(* IEC 61131-3 sources: llm-plc-st-eval/data/processed_definitivo/qwen2.5-coder_14b/B6/zero_shot, 3 files *)

(* ---- ejec_1.st ---- *)
FUNCTION_BLOCK FB_Baliza
VAR_INPUT
    alarma : BOOL;  // Variable de entrada que indica si hay una alarma
END_VAR

VAR_OUTPUT
    lampara : BOOL;  // Variable de salida que controla el estado de la lámpara
END_VAR

VAR
    timer : TON;  // Timer de conteo hacia arriba
    estado : BOOL;  // Variable para controlar el estado de parpadeo
END_VAR

// Inicialización del timer
IF timer.Q = FALSE THEN
    timer(IN := TRUE, PT := T#1S);
END_IF;

// Logica de parpadeo
IF alarma THEN
    lampara := estado;
    IF timer.Q THEN
        estado := NOT estado;  // Cambia el estado de la lámpara
        timer(IN := FALSE);  // Reinicia el timer
        timer(IN := TRUE);  // Reinicia el timer
    END_IF;
ELSE
    lampara := FALSE;  // Apaga la lámpara si no hay alarma
END_IF;

(* ---- ejec_2.st ---- *)
FUNCTION_BLOCK FB_Baliza
VAR_INPUT
    alarma : BOOL; // Variable de entrada que indica si hay una alarma
END_VAR

VAR_OUTPUT
    lampara : BOOL; // Variable de salida que controla el estado de la lámpara
END_VAR

VAR
    timer : TON; // Timer de conteo hacia arriba
    estado : BOOL; // Estado actual de la lámpara (encendida/apagada)
END_VAR

// Inicialización del timer
IF timer.Q = FALSE THEN
    timer(IN := TRUE, PT := T#1S);
END_IF;

// Lógica de la baliza
IF alarma THEN
    // Si hay alarma, la lámpara parpadea
    lampara := estado;
    IF timer.Q THEN
        // Cambia el estado de la lámpara al final del ciclo de 1 segundo
        estado := NOT estado;
        timer(IN := FALSE); // Reinicia el timer
        timer(IN := TRUE); // Reinicia el timer
    END_IF;
ELSE
    // Si no hay alarma, la lámpara permanece apagada
    lampara := FALSE;
END_IF;
END_FUNCTION_BLOCK

(* ---- ejec_3.st ---- *)
FUNCTION_BLOCK FB_Baliza
VAR_INPUT
    alarma : BOOL; // Variable de entrada que indica si hay una alarma
END_VAR

VAR_OUTPUT
    lampara : BOOL; // Variable de salida que controla el estado de la lámpara
END_VAR

VAR
    estado : BOOL := FALSE; // Variable interna para controlar el estado de parpadeo
    timer : TON; // Timer para controlar el ciclo de parpadeo
END_VAR

// Configuración del timer para un ciclo de 1 segundo
timer(IN := TRUE, PT := T#1S);

// Lógica para controlar el estado de la lámpara
IF alarma THEN
    // Si hay alarma, la lámpara parpadea
    lampara := estado;
    // Cambiar el estado de la lámpara al final del ciclo del timer
    IF timer.Q THEN
        estado := NOT estado;
        timer(IN := FALSE); // Reiniciar el timer
    END_IF
ELSE
    // Si no hay alarma, la lámpara permanece apagada
    lampara := FALSE;
END_IF
